(* IEC 61131-3 sources: llm-plc-st-eval/data/definitivo/qwen2.5-coder_14b/I4/few_shot, 3 files *)

(* ---- ejec_1.st ---- *)
FUNCTION_BLOCK FB_EstrellaTriangulo
VAR_INPUT
    btnMarcha : BOOL; (* Botón de marcha *)
    btnParo : BOOL; (* Botón de paro *)
END_VAR
VAR_OUTPUT
    kM : BOOL; (* Contactor principal *)
    kY : BOOL; (* Contactor de estrella *)
    kD : BOOL; (* Contactor de triángulo *)
END_VAR
VAR
    tEstrella : TP; (* Temporizador para el contacto de estrella *)
    tMuerto : TP; (* Temporizador para el tiempo muerto *)
    estado : INT; (* Variable de estado para el arranque estrella-triángulo *)
END_VAR

(* Estado 0: Esperando inicio *)
(* Estado 1: Contacto de estrella activo *)
(* Estado 2: Tiempo muerto *)
(* Estado 3: Contacto de triángulo activo *)

(* Botón de paro desactiva todos los contactores *)
IF btnParo THEN
    kM := FALSE;
    kY := FALSE;
    kD := FALSE;
    estado := 0;
ELSIF btnMarcha THEN
    CASE estado OF
        0:
            (* Inicia el arranque estrella-triángulo *)
            kM := TRUE;
            kY := TRUE;
            kD := FALSE;
            tEstrella(IN := TRUE, PT := T#8S);
            estado := 1;
        1:
            (* Espera el fin del temporizador de estrella *)
            IF tEstrella.Q THEN
                kY := FALSE;
                tMuerto(IN := TRUE, PT := T#100MS);
                estado := 2;
            END_IF;
        2:
            (* Espera el fin del tiempo muerto *)
            IF tMuerto.Q THEN
                kD := TRUE;
                estado := 3;
            END_IF;
        3:
            (* Mantén el contacto de triángulo activo *)
            kY := FALSE;
    END_CASE;
END_IF;
END_FUNCTION_BLOCK

(* ---- ejec_2.st ---- *)
FUNCTION_BLOCK FB_EstrellaTriangulo
VAR_INPUT
    btnMarcha : BOOL; (* Boton de marcha *)
    btnParo : BOOL; (* Boton de paro *)
END_VAR
VAR_OUTPUT
    kM : BOOL; (* Contactor principal *)
    kY : BOOL; (* Contactor de estrella *)
    kD : BOOL; (* Contactor de triangulo *)
END_VAR
VAR
    tEstrella : TP; (* Temporizador para el contacto de estrella *)
    tMuerto : TP; (* Temporizador para el tiempo muerto *)
    estado : INT := 0; (* Estado actual del arranque *)
END_VAR

(* Estado 0: Esperando el botón de marcha *)
IF btnMarcha AND estado = 0 THEN
    estado := 1;
    kM := TRUE;
    kY := TRUE;
    kD := FALSE;
    tEstrella(IN := TRUE, PT := T#8S);
ELSIF btnParo THEN
    estado := 0;
    kM := FALSE;
    kY := FALSE;
    kD := FALSE;
END_IF

(* Estado 1: Esperando el temporizador de estrella *)
IF estado = 1 AND tEstrella.Q THEN
    estado := 2;
    kY := FALSE;
    tMuerto(IN := TRUE, PT := T#100MS);
END_IF

(* Estado 2: Esperando el tiempo muerto *)
IF estado = 2 AND tMuerto.Q THEN
    estado := 3;
    kD := TRUE;
END_IF

(* Mantener kY y kD inactivos simultáneamente *)
IF kY AND kD THEN
    kY := FALSE;
    kD := FALSE;
END_IF

END_FUNCTION_BLOCK

(* ---- ejec_3.st ---- *)
FUNCTION_BLOCK FB_EstrellaTriangulo
VAR_INPUT
    btnMarcha : BOOL; (* Botón de marcha *)
    btnParo : BOOL; (* Botón de paro *)
END_VAR
VAR_OUTPUT
    kM : BOOL; (* Contactor principal *)
    kY : BOOL; (* Contactor de estrella *)
    kD : BOOL; (* Contactor de triángulo *)
END_VAR
VAR
    tEstrella : TP; (* Temporizador para el contacto de estrella *)
    tMuerto : TP; (* Temporizador para el tiempo muerto *)
    estado : INT; (* Estado actual del arranque estrella-triángulo *)
END_VAR

(* Estados del arranque estrella-triángulo *)
CONST
    ESTADO_INICIAL := 0;
    ESTADO_ESTRELLA := 1;
    ESTADO_MUERTO := 2;
    ESTADO_TRIANGULO := 3;
END_CONST

(* Paro inmediato *)
IF btnParo THEN
    kM := FALSE;
    kY := FALSE;
    kD := FALSE;
    estado := ESTADO_INICIAL;
ELSIF btnMarcha THEN
    CASE estado OF
        ESTADO_INICIAL:
            kM := TRUE;
            kY := TRUE;
            kD := FALSE;
            tEstrella(IN := TRUE, PT := T#8S);
            estado := ESTADO_ESTRELLA;
        ESTADO_ESTRELLA:
            IF tEstrella.Q THEN
                kY := FALSE;
                tMuerto(IN := TRUE, PT := T#100MS);
                estado := ESTADO_MUERTO;
            END_IF;
        ESTADO_MUERTO:
            IF tMuerto.Q THEN
                kD := TRUE;
                estado := ESTADO_TRIANGULO;
            END_IF;
        ESTADO_TRIANGULO:
            (* Mantener kD activo mientras kY esté inactivo *)
            kD := TRUE;
    END_CASE;
END_IF;

(* Asegurar que kY y kD no estén activos simultáneamente *)
IF kY AND kD THEN
    kY := FALSE;
END_IF;

END_FUNCTION_BLOCK
